TYPE ST_CamMasterParam :
STRUCT
	fMasterFactor: LREAL;
	fMasterVelo: LREAL;
	fMasterAngeleMax: LREAL;
	fMasterAngeleMin: LREAL;
END_STRUCT
END_TYPE

(* stored: Version 1.1.0.1, ProductVersion 3.1.4024.12
   DUT ST_CamMasterParam: Id {914ac56b-87d1-46c3-8ccf-c1cdf7b0c3c6} *)
